// TwinCAT 3 PLC project TestPLC
// ProgramVersion: 3.1.4026.27
// libraries:
//   PersistentDataHandler, * (Beckhoff Community)
//   Tc2_Standard, * (Beckhoff Automation GmbH)
//   Tc2_System, * (Beckhoff Automation GmbH)
// project tree:
//   GVLs/ GVL.TcGVL
//   / PersistentTask.TcTTO, PlcTask.TcTTO
//   POUs/ FB_Example.TcPOU, MAIN.TcPOU, PersistentCaller.TcPOU
// (motion and I/O tree: see PLC project persistentdatahandler)
// real-time tasks:
//   TASK PlcTask: cycle T#10ms, priority 20, ADS port 350
//   TASK PersistentTask: cycle T#200us, priority 1, ADS port 351
// variable links:

CONFIGURATION TestPLC
    RESOURCE PLC ON TwinCAT3
        TASK PersistentTask(INTERVAL := T#200us, PRIORITY := 1);
        TASK PlcTask(INTERVAL := T#10ms, PRIORITY := 20);
        PROGRAM PersistentCaller WITH PersistentTask : PersistentCaller;
        PROGRAM MAIN WITH PlcTask : MAIN;
    END_RESOURCE
END_CONFIGURATION

// ---- GVLs/GVL.TcGVL
{attribute 'qualified_only'}
VAR_GLOBAL PERSISTENT
	persist_int 	: INT;
	persist_str 	: T_MaxString;
	persist_float	: REAL;
END_VAR

// ---- POUs/PersistentCaller.TcPOU
PROGRAM PersistentCaller
VAR
	persistanceHandler : FB_PersistentHandler;
	enable	: BOOL := TRUE;
	reinit	: BOOL := FALSE;
END_VAR


persistanceHandler(bEnable := enable,
				   bReinit := reinit);

END_PROGRAM

// ---- POUs/MAIN.TcPOU
PROGRAM MAIN
VAR
	example : FB_Example;
	filler : ARRAY[0..130] OF FB_Example;
	
	wroteData : BOOL;
	loadedData : BOOL;
END_VAR
VAR PERSISTENT
	per_example : FB_Example;
END_VAR

END_PROGRAM

// ---- POUs/FB_Example.TcPOU
FUNCTION_BLOCK FB_Example
VAR PERSISTENT
	persist_int 	: INT;
	persist_str 	: T_MaxString;
	persist_float	: REAL;
END_VAR
VAR RETAIN
	retain_int 		: INT;
	retain_str 		: T_MaxString;
	retain_float	: REAL;
END_VAR
VAR 
	non_per		: INT;
	non_per2	: LREAL;
	timer		: TON;
END_VAR

END_FUNCTION_BLOCK
